// TIA Portal V20 export
Screen "190RB02_J5"  1276x673
  ScreenItem "Line_Header_X0_Y64" at 0,64 size 1276x0  Type=HmiLine
  ScreenItem "permanentareaborderrectangle" at 0,0 size 0x0  Type=HmiRectangle
  ScreenItem "Button_Back" at 2,2 size 90x60  Type=HmiButton
  ScreenItem "Title_ScreenOverview_X390_Y2_1" at 390,3 size 510x57  Type=HmiTextBox
  ScreenItem "Fusszeile_Button_ManualOPMode1_4" at 1181,2 size 90x60  Type=HmiButton
  ScreenItem "Graphic view_1" at 195,100 size 801x526  Type=HmiGraphicView
  ScreenItem "Line_4" at 630,166 size 56x114  Type=HmiLine
  ScreenItem "Fusszeile_Button_ManualOPMode1_1" at 1088,2 size 90x60  Type=HmiButton
  ScreenItem "Title_ScreenOverview_X390_Y2_5" at 1130,78 size 139x57  Type=HmiTextBox
  ScreenItem "Title_ScreenOverview_X390_Y2_6" at 1130,144 size 139x57  Type=HmiTextBox
  ScreenItem "Title_ScreenOverview_X390_Y2_7" at 1130,144 size 139x57  Type=HmiTextBox
  ScreenItem "文本域_1" at 900,72 size 134x40  Type=HmiTextBox
  ScreenItem "Line_3" at 844,134 size 76x144  Type=HmiLine
  ScreenItem "Line_10" at 872,213 size 91x71  Type=HmiLine
  ScreenItem "文本域_2" at 1031,240 size 134x40  Type=HmiTextBox
  ScreenItem "Line_11" at 949,262 size 77x1  Type=HmiLine
  ScreenItem "文本域_5" at 1130,294 size 134x40  Type=HmiTextBox
  ScreenItem "Line_12" at 944,288 size 206x68  Type=HmiLine
  ScreenItem "文本域_6" at 1059,377 size 134x40  Type=HmiTextBox
  ScreenItem "Line_13" at 864,365 size 186x31  Type=HmiLine
  ScreenItem "文本域_7" at 1136,467 size 134x40  Type=HmiTextBox
  ScreenItem "Line_14" at 942,445 size 185x41  Type=HmiLine
  ScreenItem "文本域_8" at 1103,567 size 134x40  Type=HmiTextBox
  ScreenItem "Line_15" at 853,444 size 241x117  Type=HmiLine
  ScreenItem "文本域_3" at 916,567 size 134x40  Type=HmiTextBox
  ScreenItem "Line_1" at 700,360 size 221x196  Type=HmiLine
  ScreenItem "Line_2" at 637,456 size 71x97  Type=HmiLine
  ScreenItem "文本域_4" at 650,567 size 134x40  Type=HmiTextBox
  ScreenItem "Line_5" at 440,456 size 15x107  Type=HmiLine
  ScreenItem "文本域_9" at 390,567 size 134x40  Type=HmiTextBox
  ScreenItem "Line_6" at 304,411 size 53x151  Type=HmiLine
  ScreenItem "文本域_10" at 232,567 size 134x40  Type=HmiTextBox
  ScreenItem "Line_7" at 147,443 size 148x124  Type=HmiLine
  ScreenItem "文本域_12" at 64,570 size 134x40  Type=HmiTextBox
  ScreenItem "文本域_13" at 17,405 size 134x40  Type=HmiTextBox
  ScreenItem "Line_8" at 159,424 size 73x13  Type=HmiLine
  ScreenItem "Line_9" at 169,340 size 123x56  Type=HmiLine
  ScreenItem "Line_16" at 496,154 size 54x103  Type=HmiLine
  ScreenItem "文本域_16" at 31,201 size 134x40  Type=HmiTextBox
  ScreenItem "Line_17" at 173,233 size 73x63  Type=HmiLine
  ScreenItem "文本域_17" at 70,96 size 134x40  Type=HmiTextBox
  ScreenItem "Line_18" at 212,128 size 148x188  Type=HmiLine
  ScreenItem "文本域_18" at 247,76 size 134x40  Type=HmiTextBox
  ScreenItem "Line_19" at 342,128 size 91x142  Type=HmiLine
  ScreenItem "Rectangle_13" at 0,0 size 152x48  Type=HmiRectangle
  ScreenItem "文本域_19" at 2,1 size 122x45  Type=HmiTextBox
  ScreenItem "圆_5" at 0,0 size 100x30  Type=HmiCircle
  ScreenItem "圆_6" at 0,0 size 100x30  Type=HmiCircle
  ScreenItem "Title_ScreenOverview_X390_Y2_4" at 689,164 size 52x19  Type=HmiTextBox
  ScreenItem "Title_ScreenOverview_X390_Y2_3" at 716,184 size 25x21  Type=HmiTextBox
  ScreenItem "Title_ScreenOverview_X390_Y2_2" at 689,184 size 25x21  Type=HmiTextBox
  ScreenItem "文本域_15" at 648,120 size 134x40  Type=HmiTextBox
  ScreenItem "Title_ScreenOverview_X390_Y2_8" at 930,112 size 52x19  Type=HmiTextBox
  ScreenItem "Title_ScreenOverview_X390_Y2_9" at 957,132 size 25x21  Type=HmiTextBox
  ScreenItem "Title_ScreenOverview_X390_Y2_10" at 930,132 size 25x21  Type=HmiTextBox
  ScreenItem "Title_ScreenOverview_X390_Y2_11" at 1059,278 size 52x19  Type=HmiTextBox
  ScreenItem "Title_ScreenOverview_X390_Y2_12" at 1059,298 size 25x21  Type=HmiTextBox
  ScreenItem "Title_ScreenOverview_X390_Y2_13" at 1086,298 size 25x21  Type=HmiTextBox
  ScreenItem "Title_ScreenOverview_X390_Y2_14" at 1162,336 size 52x19  Type=HmiTextBox
  ScreenItem "Title_ScreenOverview_X390_Y2_15" at 1162,356 size 25x21  Type=HmiTextBox
  ScreenItem "Title_ScreenOverview_X390_Y2_16" at 1189,356 size 25x21  Type=HmiTextBox
  ScreenItem "Title_ScreenOverview_X390_Y2_17" at 1106,417 size 52x19  Type=HmiTextBox
  ScreenItem "Title_ScreenOverview_X390_Y2_18" at 1106,437 size 25x21  Type=HmiTextBox
  ScreenItem "Title_ScreenOverview_X390_Y2_19" at 1133,437 size 25x21  Type=HmiTextBox
  ScreenItem "Title_ScreenOverview_X390_Y2_20" at 1168,508 size 52x19  Type=HmiTextBox
  ScreenItem "Title_ScreenOverview_X390_Y2_21" at 1168,528 size 25x21  Type=HmiTextBox
  ScreenItem "Title_ScreenOverview_X390_Y2_22" at 1195,528 size 25x21  Type=HmiTextBox
  ScreenItem "Title_ScreenOverview_X390_Y2_23" at 1150,607 size 52x19  Type=HmiTextBox
  ScreenItem "Title_ScreenOverview_X390_Y2_24" at 1150,627 size 25x21  Type=HmiTextBox
  ScreenItem "Title_ScreenOverview_X390_Y2_25" at 1177,627 size 25x21  Type=HmiTextBox
  ScreenItem "Title_ScreenOverview_X390_Y2_26" at 990,629 size 25x21  Type=HmiTextBox
  ScreenItem "Title_ScreenOverview_X390_Y2_27" at 963,609 size 52x19  Type=HmiTextBox
  ScreenItem "Title_ScreenOverview_X390_Y2_28" at 963,629 size 25x21  Type=HmiTextBox
  ScreenItem "Title_ScreenOverview_X390_Y2_29" at 713,629 size 25x21  Type=HmiTextBox
  ScreenItem "Title_ScreenOverview_X390_Y2_30" at 686,609 size 52x19  Type=HmiTextBox
  ScreenItem "Title_ScreenOverview_X390_Y2_31" at 686,629 size 25x21  Type=HmiTextBox
  ScreenItem "Title_ScreenOverview_X390_Y2_32" at 282,610 size 52x19  Type=HmiTextBox
  ScreenItem "Title_ScreenOverview_X390_Y2_33" at 282,630 size 25x21  Type=HmiTextBox
  ScreenItem "Title_ScreenOverview_X390_Y2_34" at 309,630 size 25x21  Type=HmiTextBox
  ScreenItem "Title_ScreenOverview_X390_Y2_35" at 433,610 size 52x19  Type=HmiTextBox
  ScreenItem "Title_ScreenOverview_X390_Y2_36" at 433,630 size 25x21  Type=HmiTextBox
  ScreenItem "Title_ScreenOverview_X390_Y2_37" at 460,630 size 25x21  Type=HmiTextBox
  ScreenItem "Title_ScreenOverview_X390_Y2_38" at 107,611 size 52x19  Type=HmiTextBox
  ScreenItem "Title_ScreenOverview_X390_Y2_39" at 107,631 size 25x21  Type=HmiTextBox
  ScreenItem "Title_ScreenOverview_X390_Y2_40" at 134,631 size 25x21  Type=HmiTextBox
  ScreenItem "Title_ScreenOverview_X390_Y2_41" at 47,445 size 52x19  Type=HmiTextBox
  ScreenItem "Title_ScreenOverview_X390_Y2_42" at 47,465 size 25x21  Type=HmiTextBox
  ScreenItem "Title_ScreenOverview_X390_Y2_43" at 74,465 size 25x21  Type=HmiTextBox
  ScreenItem "Title_ScreenOverview_X390_Y2_44" at 74,244 size 52x19  Type=HmiTextBox
  ScreenItem "Title_ScreenOverview_X390_Y2_45" at 74,264 size 25x21  Type=HmiTextBox
  ScreenItem "Title_ScreenOverview_X390_Y2_46" at 101,264 size 25x21  Type=HmiTextBox
  ScreenItem "Title_ScreenOverview_X390_Y2_47" at 112,139 size 52x19  Type=HmiTextBox
  ScreenItem "Title_ScreenOverview_X390_Y2_48" at 112,159 size 25x21  Type=HmiTextBox
  ScreenItem "Title_ScreenOverview_X390_Y2_49" at 139,159 size 25x21  Type=HmiTextBox
  ScreenItem "Title_ScreenOverview_X390_Y2_50" at 280,118 size 52x19  Type=HmiTextBox
  ScreenItem "Title_ScreenOverview_X390_Y2_51" at 280,138 size 25x21  Type=HmiTextBox
  ScreenItem "Title_ScreenOverview_X390_Y2_52" at 307,138 size 25x21  Type=HmiTextBox
  ScreenItem "Rectangle_1" at 0,0 size 152x48  Type=HmiRectangle
  ScreenItem "文本域_11" at 2,1 size 122x45  Type=HmiTextBox
  ScreenItem "圆_1" at 0,0 size 100x30  Type=HmiCircle
  ScreenItem "圆_2" at 0,0 size 100x30  Type=HmiCircle
  ScreenItem "Rectangle_2" at 0,0 size 152x48  Type=HmiRectangle
  ScreenItem "文本域_14" at 2,1 size 122x45  Type=HmiTextBox
  ScreenItem "圆_3" at 0,0 size 100x30  Type=HmiCircle
  ScreenItem "圆_4" at 0,0 size 100x30  Type=HmiCircle
